(* IEC 61131-3 sources: llm-plc-st-eval/data/definitivo/qwen2.5-coder_14b/C7/zero_shot, 3 files *)

(* ---- ejec_1.st ---- *)
```pascal
FUNCTION_BLOCK FB_Contador
VAR_INPUT
    sensorPieza : BOOL; // Contacto normalmente abierto sensor de pieza
    btnReset : BOOL;    // Contacto normalmente abierto botón de reset
END_VAR

VAR_OUTPUT
    loteListo : BOOL; // Bobina que indica que el lote está listo
    cuenta : INT;      // Variable que almacena el valor actual del contador
END_VAR

VAR
    C1 : CTU;          // Contador ascendente
END_VAR

// Configuración del contador C1
C1.PV := 12;          // Valor preestablecido del contador

// Rama 1: Conteo de piezas
C1(CU := sensorPieza, RESET := btnReset);

// Rama 2: Indicación de lote listo
loteListo := C1.Q;

// Rama 3: Transferencia del valor actual del contador a la variable cuenta
cuenta := C1.CV;
END_FUNCTION_BLOCK
```

Este código en Structured Text (ST) implementa el comportamiento descrito en el Ladder Diagram, utilizando un FUNCTION_BLOCK llamado `FB_Contador` con las variables de entrada y salida especificadas. El contador ascendente `C1` se configura con un valor preestablecido de 12, y las ramas del programa se implementan según la descripción proporcionada.

(* ---- ejec_2.st ---- *)
```pascal
FUNCTION_BLOCK FB_Contador
VAR_INPUT
    sensorPieza : BOOL; // Contacto normalmente abierto del sensor de pieza
    btnReset : BOOL;    // Contacto normalmente abierto del botón de reset
END_VAR

VAR_OUTPUT
    loteListo : BOOL;  // Bobina que indica que el lote está listo
    cuenta : INT;      // Variable que almacena el valor actual del contador
END_VAR

VAR
    C1 : CTU;          // Contador ascendente
END_VAR

// Configuración del contador ascendente
C1.PV := 12;          // Valor preestablecido del contador

// Rama 1: Conteo de piezas
C1(CU := sensorPieza, RESET := btnReset);

// Rama 2: Indicación de lote listo
loteListo := C1.Q;

// Rama 3: Transferencia del valor actual del contador a la variable cuenta
cuenta := C1.CV;
END_FUNCTION_BLOCK
```

(* ---- ejec_3.st ---- *)
```pascal
FUNCTION_BLOCK FB_Contador
VAR_INPUT
    sensorPieza : BOOL; // Contacto normalmente abierto sensor de pieza
    btnReset : BOOL; // Contacto normalmente abierto botón de reset
END_VAR

VAR_OUTPUT
    loteListo : BOOL; // Bobina que indica que el lote está listo
    cuenta : INT; // Variable que almacena el valor actual del contador
END_VAR

VAR
    C1 : CTU; // Contador ascendente
END_VAR

// Configuración del contador ascendente
C1.PV := 12; // Valor preestablecido del contador

// Rama 1: Conteo de piezas
IF sensorPieza THEN
    C1.CU := TRUE; // Alimenta la entrada de conteo
ELSE
    C1.CU := FALSE;
END_IF;

// Rama 2: Reset del contador
IF btnReset THEN
    C1.RESET := TRUE; // Alimenta la entrada de reset
ELSE
    C1.RESET := FALSE;
END_IF;

// Rama 3: Transferencia del valor del contador a la variable cuenta
cuenta := C1.CV; // Transfiere el valor actual del contador a la variable cuenta

// Rama 4: Control de la bobina loteListo
IF C1.Q THEN
    loteListo := TRUE; // Activa la bobina si el contador alcanza el valor preestablecido
ELSE
    loteListo := FALSE;
END_IF;

END_FUNCTION_BLOCK
```
